TYPE ST_MBSignalConfig :
STRUCT
    modbusAddr          : UDINT;
    dataType            : E_MBDataType;
    bitIndex            : BYTE := 255;
    tag                 : STRING(32);
END_STRUCT
END_TYPE

(* stored: Version 1.1.0.1, ProductVersion 3.1.4024.0
   DUT ST_MBSignalConfig: Id {8b1cdb32-47f9-48c3-88c0-6adde8ce65ca} *)
